# EPICS substitutions: db/Beckhoff_7XXX/ecmcEP7211-0034_OPT_info2Temp.substitutions
file "ecmc_analogInput-chX.template"
{
  pattern {CH_ID, sourceName, KEY,   suffix,    DESC,        EGU,    ESLO, PREC, LOPR, HOPR, LOLO, LOW, HIGH, HIHI, HYST, LLSV,       LSV,        HSV,     HHSV}
          {02,    "infoData", "Drv", "-TmpAct", "InfoData2", "degC", 0.1,  1,    0,    50,   0,    0,   40,   50,   0.5,  "NO_ALARM", "NO_ALARM", "MINOR", "MAJOR"}
}
